(* IEC 61131-3 sources: s7-to-codesys/tests/POUs/S7Compat/FB_S5Timer_Test, 9 files *)

(* ---- BcdCarriesTimeBase.method.decl.st ---- *)
// SD, S5T#20S: шкала 100 мс, 200 единиц; LC T — BCD со шкалой (16#1200, через 5 с — 16#1150); L T
// округляет остаток вверх (через 5050 мс — 150 единиц).
METHOD PRIVATE BcdCarriesTimeBase
VAR
    stTimer : ST_S5Timer;   // проверяемый таймер
    wPreset : WORD;         // S5T#20S
END_VAR

(* ---- EnableRestartsRunningTimer.method.decl.st ---- *)
// FR + SE, S5T#1S: фронт FR при RLO пуска = 1 перезапускает идущий таймер; спад FR ничего не делает; новый
// фронт FR снова даёт пуск без фронта RLO пуска (AWL_e.pdf §12.3).
METHOD PRIVATE EnableRestartsRunningTimer
VAR
    stTimer : ST_S5Timer;   // проверяемый таймер
    wPreset : WORD;         // S5T#1S
END_VAR

(* ---- ExtPulseRunsOutAndRetriggers.method.decl.st ---- *)
// SE, S5T#1S: Q держится после спада RLO; фронт на 600 мс перезапускает таймер — истечение на 1600 мс.
METHOD PRIVATE ExtPulseRunsOutAndRetriggers
VAR
    stTimer : ST_S5Timer;   // проверяемый таймер
    wPreset : WORD;         // S5T#1S
END_VAR

(* ---- OffDelayHoldsAfterFall.method.decl.st ---- *)
// SF, S5T#1S: Q = TRUE при RLO = 1 и 1000 мс после спада; фронт RLO останавливает идущий таймер (остаток
// 50 единиц), следующий спад запускает его заново.
METHOD PRIVATE OffDelayHoldsAfterFall
VAR
    stTimer : ST_S5Timer;   // проверяемый таймер
    wPreset : WORD;         // S5T#1S
END_VAR

(* ---- OnDelayNeedsRloHeld.method.decl.st ---- *)
// SD, S5T#1S: Q = TRUE ровно через 1000 мс при RLO = 1; RLO = 0 сбрасывает Q и останавливает таймер с
// остатком (70 единиц через 300 мс после повторного пуска) — и через 1 с остаток тот же, Q = FALSE.
METHOD PRIVATE OnDelayNeedsRloHeld
VAR
    stTimer : ST_S5Timer;   // проверяемый таймер
    wPreset : WORD;         // S5T#1S
END_VAR

(* ---- PulseStopsWhenRloFalls.method.decl.st ---- *)
// SP, S5T#1S (шкала 10 мс): Q, пока таймер идёт и RLO = 1; по истечении Q = FALSE без перезапуска; RLO = 0
// останавливает таймер, остаток сохраняется (90 единиц через 100 мс после пуска).
METHOD PRIVATE PulseStopsWhenRloFalls
VAR
    stTimer : ST_S5Timer;   // проверяемый таймер (новый на каждый вызов метода)
    wPreset : WORD;         // S5T#1S
END_VAR

(* ---- QReadBeforeStartSeesPreviousState.method.decl.st ---- *)
// Опрос до инструкции пуска в том же цикле: SD, S5T#1S, на 1000 мс время истекло — чтение до SD видит
// Q = TRUE, SD с RLO = 0 сбрасывает Q, чтение после — FALSE. В S7 таймер обновляет часовой процесс CPU, и
// опрос из любого места программы видит одно и то же слово таймера (GVL_S5Timers — общий для всех блоков).
METHOD PRIVATE QReadBeforeStartSeesPreviousState
VAR
    stTimer : ST_S5Timer;   // проверяемый таймер
    wPreset : WORD;         // S5T#1S
END_VAR

(* ---- ResetIsLevelAndNeedsNewEdge.method.decl.st ---- *)
// SD + R, S5T#1S: R при RLO = 1 держит таймер сброшенным; после снятия сброса без нового фронта пуска таймер
// не идёт (Q = FALSE и через 2 с), новый фронт запускает его.
METHOD PRIVATE ResetIsLevelAndNeedsNewEdge
VAR
    stTimer : ST_S5Timer;   // проверяемый таймер
    wPreset : WORD;         // S5T#1S
END_VAR

(* ---- RetOnDelayHoldsQUntilReset.method.decl.st ---- *)
// SS, S5T#1S: время истекает и при RLO = 0, Q = TRUE держится до R; после сброса — новый пуск фронтом.
METHOD PRIVATE RetOnDelayHoldsQUntilReset
VAR
    stTimer : ST_S5Timer;   // проверяемый таймер
    wPreset : WORD;         // S5T#1S
END_VAR
